FUNCTION_BLOCK Distributing (* CAT Function Block Type *)
  (* Standard: 61499-2 *)
  (* Version 0.0, 11/16/2026, Sandeep Patil, Flexbridge AB, template *)
  PACKAGE Flexbridge.FestoMPS400;
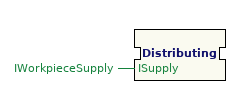
  SOCKETS
    ISupply : IWorkpieceSupply;
  END_SOCKETS
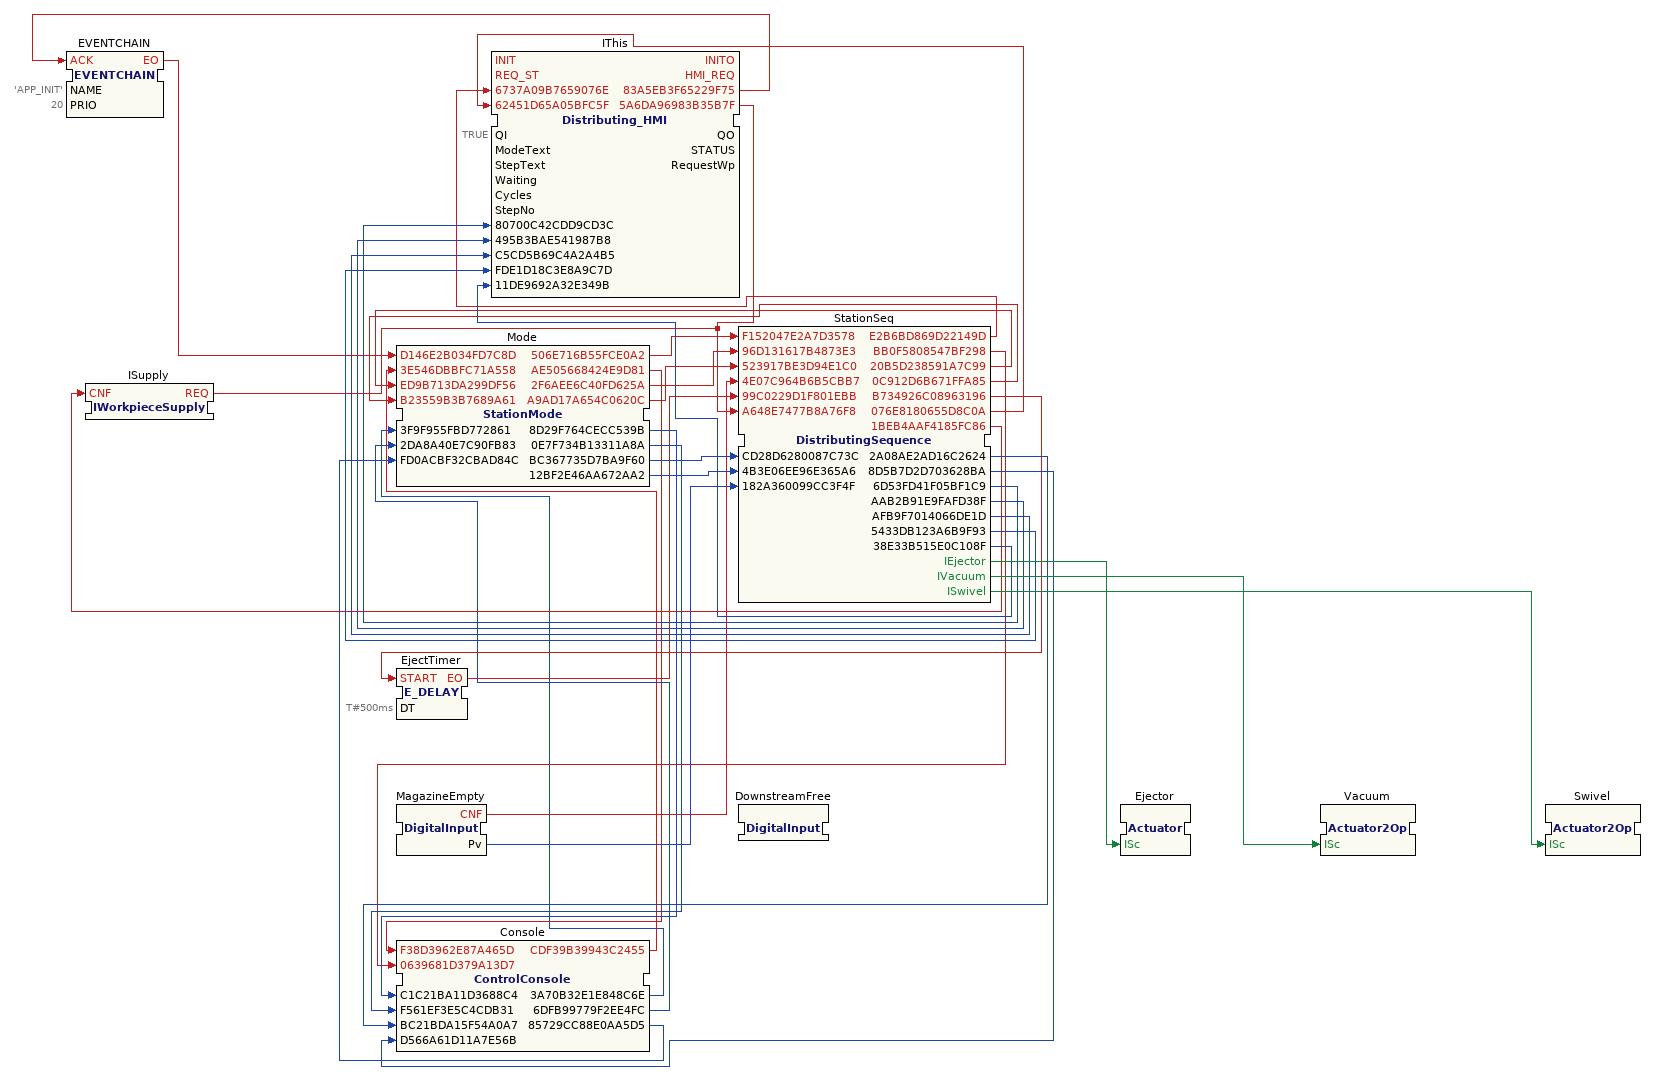
  (* 0 - INITIALIZATION *)
  (* 6 - HMI INTERFACE *)
  (* 1 - FUNCTIONAL INPUT INTERFACE *)
  (* 5 - LOGICS *)
  (* 2 - FUNCTIONAL OUTPUT INTERFACE *)
  (* 3 - FIELD INTERFACE (3.B FROM THE FIELD: plain sensors) *)
  (* 4 - CHILDREN *)
  (* 4.A - TYPICALS (one device CAT per Festo device) *)
  FBS
    Ejector : Actuator;
    Vacuum : Actuator2Op;
    Swivel : Actuator2Op;
    MagazineEmpty : DigitalInput;
    DownstreamFree : DigitalInput;
    EVENTCHAIN : EVENTCHAIN(NAME := 'APP_INIT', PRIO := 20);
    IThis : Distributing_HMI(QI := TRUE);
    Mode : StationMode;
    StationSeq : DistributingSequence;
    EjectTimer : E_DELAY(DT := T#500ms);
    Console : ControlConsole;
  END_FBS
  EVENT_CONNECTIONS
    EVENTCHAIN.EO TO Mode.D146E2B034FD7C8D;
    Mode.506E716B55FCE0A2 TO StationSeq.F152047E2A7D3578;
    StationSeq.E2B6BD869D22149D TO IThis.6737A09B7659076E;
    IThis.83A5EB3F65229F75 TO EVENTCHAIN.ACK;
    Console.CDF39B39943C2455 TO Mode.3E546DBBFC71A558;
    Mode.AE505668424E9D81 TO Console.F38D3962E87A465D;
    StationSeq.BB0F5808547BF298 TO Console.0639681D379A13D7;
    Mode.2F6AEE6C40FD625A TO StationSeq.96D131617B4873E3;
    StationSeq.20B5D238591A7C99 TO Mode.ED9B713DA299DF56;
    StationSeq.0C912D6B671FFA85 TO Mode.B23559B3B7689A61;
    Mode.A9AD17A654C0620C TO StationSeq.523917BE3D94E1C0;
    MagazineEmpty.CNF TO StationSeq.4E07C964B6B5CBB7;
    StationSeq.B734926C08963196 TO EjectTimer.START;
    EjectTimer.EO TO StationSeq.99C0229D1F801EBB;
    StationSeq.076E8180655D8C0A TO IThis.62451D65A05BFC5F;
    IThis.5A6DA96983B35B7F TO StationSeq.A648E7477B8A76F8;
    ISupply.REQ TO StationSeq.A648E7477B8A76F8;
    StationSeq.1BEB4AAF4185FC86 TO ISupply.CNF;
  END_CONNECTIONS
  DATA_CONNECTIONS
    Console.3A70B32E1E848C6E TO Mode.3F9F955FBD772861;
    Console.6DFB99779F2EE4FC TO Mode.2DA8A40E7C90FB83;
    Console.85729CC88E0AA5D5 TO Mode.FD0ACBF32CBAD84C;
    Mode.8D29F764CECC539B TO Console.C1C21BA11D3688C4;
    Mode.0E7F734B13311A8A TO Console.F561EF3E5C4CDB31;
    StationSeq.2A08AE2AD16C2624 TO Console.BC21BDA15F54A0A7;
    StationSeq.8D5B7D2D703628BA TO Console.D566A61D11A7E56B;
    Mode.BC367735D7BA9F60 TO StationSeq.CD28D6280087C73C;
    Mode.12BF2E46AA672AA2 TO StationSeq.4B3E06EE96E365A6;
    MagazineEmpty.Pv TO StationSeq.182A360099CC3F4F;
    StationSeq.6D53FD41F05BF1C9 TO IThis.80700C42CDD9CD3C;
    StationSeq.AAB2B91E9FAFD38F TO IThis.495B3BAE541987B8;
    StationSeq.AFB9F7014066DE1D TO IThis.C5CD5B69C4A2A4B5;
    StationSeq.5433DB123A6B9F93 TO IThis.FDE1D18C3E8A9C7D;
    StationSeq.38E33B515E0C108F TO IThis.11DE9692A32E349B;
  END_CONNECTIONS
  ADAPTER_CONNECTIONS
    StationSeq.IEjector TO Ejector.ISc;
    StationSeq.IVacuum TO Vacuum.ISc;
    StationSeq.ISwivel TO Swivel.ISc;
  END_CONNECTIONS
END_FUNCTION_BLOCK
